// TIA Portal V18 export
TYPE "UserValidationMdz_out"
   STRUCT
      Station : Array[1.."Station_Setup_Const"] of Struct
         Position : Array[1.."Position_Setup_Const"] of Struct
            User_ID : DInt;
            User_SSB : String[8];
            UserName : String[37];
            MsgLogin : String[40];
            AuthorizedByUserMaster_ID : DInt;
            Authentication : Bool;
         END_STRUCT;
      END_STRUCT;
   END_STRUCT;
   // Station[1].Position[1].User_ID := 0;
   // Station[2].Position[1].User_ID := 0;
   // Station[3].Position[1].User_ID := 0;
   // Station[4].Position[1].User_ID := 0;
   // Station[5].Position[1].User_ID := 0;
   // Station[6].Position[1].User_ID := 0;
   // Station[7].Position[1].User_ID := 0;
   // Station[8].Position[1].User_ID := 0;
   // Station[9].Position[1].User_ID := 0;
   // Station[10].Position[1].User_ID := 0;
   // Station[11].Position[1].User_ID := 0;
   // Station[12].Position[1].User_ID := 0;
   // Station[13].Position[1].User_ID := 0;
   // Station[14].Position[1].User_ID := 0;
   // Station[15].Position[1].User_ID := 0;
   // Station[16].Position[1].User_ID := 0;
   // Station[17].Position[1].User_ID := 0;
   // Station[18].Position[1].User_ID := 0;
   // Station[19].Position[1].User_ID := 0;
   // Station[20].Position[1].User_ID := 0;
   // Station[1].Position[1].User_SSB := '';
   // Station[2].Position[1].User_SSB := '';
   // Station[3].Position[1].User_SSB := '';
   // Station[4].Position[1].User_SSB := '';
   // Station[5].Position[1].User_SSB := '';
   // Station[6].Position[1].User_SSB := '';
   // Station[7].Position[1].User_SSB := '';
   // Station[8].Position[1].User_SSB := '';
   // Station[9].Position[1].User_SSB := '';
   // Station[10].Position[1].User_SSB := '';
   // Station[11].Position[1].User_SSB := '';
   // Station[12].Position[1].User_SSB := '';
   // Station[13].Position[1].User_SSB := '';
   // Station[14].Position[1].User_SSB := '';
   // Station[15].Position[1].User_SSB := '';
   // Station[16].Position[1].User_SSB := '';
   // Station[17].Position[1].User_SSB := '';
   // Station[18].Position[1].User_SSB := '';
   // Station[19].Position[1].User_SSB := '';
   // Station[20].Position[1].User_SSB := '';
   // Station[1].Position[1].UserName := '';
   // Station[2].Position[1].UserName := '';
   // Station[3].Position[1].UserName := '';
   // Station[4].Position[1].UserName := '';
   // Station[5].Position[1].UserName := '';
   // Station[6].Position[1].UserName := '';
   // Station[7].Position[1].UserName := '';
   // Station[8].Position[1].UserName := '';
   // Station[9].Position[1].UserName := '';
   // Station[10].Position[1].UserName := '';
   // Station[11].Position[1].UserName := '';
   // Station[12].Position[1].UserName := '';
   // Station[13].Position[1].UserName := '';
   // Station[14].Position[1].UserName := '';
   // Station[15].Position[1].UserName := '';
   // Station[16].Position[1].UserName := '';
   // Station[17].Position[1].UserName := '';
   // Station[18].Position[1].UserName := '';
   // Station[19].Position[1].UserName := '';
   // Station[20].Position[1].UserName := '';
   // Station[1].Position[1].MsgLogin := 'POSTO: 1 NAO POSSUI USUARIO CADASTRADO';
   // Station[2].Position[1].MsgLogin := 'POSTO: 1 NAO POSSUI USUARIO CADASTRADO';
   // Station[3].Position[1].MsgLogin := 'POSTO: 1 NAO POSSUI USUARIO CADASTRADO';
   // Station[4].Position[1].MsgLogin := 'POSTO: 1 NAO POSSUI USUARIO CADASTRADO';
   // Station[5].Position[1].MsgLogin := 'POSTO: 1 NAO POSSUI USUARIO CADASTRADO';
   // Station[6].Position[1].MsgLogin := 'POSTO: 1 NAO POSSUI USUARIO CADASTRADO';
   // Station[7].Position[1].MsgLogin := 'POSTO: 1 NAO POSSUI USUARIO CADASTRADO';
   // Station[8].Position[1].MsgLogin := 'POSTO: 1 NAO POSSUI USUARIO CADASTRADO';
   // Station[9].Position[1].MsgLogin := 'POSTO: 1 NAO POSSUI USUARIO CADASTRADO';
   // Station[10].Position[1].MsgLogin := 'POSTO: 1 NAO POSSUI USUARIO CADASTRADO';
   // Station[11].Position[1].MsgLogin := 'POSTO: 1 NAO POSSUI USUARIO CADASTRADO';
   // Station[12].Position[1].MsgLogin := 'POSTO: 1 NAO POSSUI USUARIO CADASTRADO';
   // Station[13].Position[1].MsgLogin := 'POSTO: 1 NAO POSSUI USUARIO CADASTRADO';
   // Station[14].Position[1].MsgLogin := 'POSTO: 1 NAO POSSUI USUARIO CADASTRADO';
   // Station[15].Position[1].MsgLogin := 'POSTO: 1 NAO POSSUI USUARIO CADASTRADO';
   // Station[16].Position[1].MsgLogin := 'POSTO: 1 NAO POSSUI USUARIO CADASTRADO';
   // Station[17].Position[1].MsgLogin := 'POSTO: 1 NAO POSSUI USUARIO CADASTRADO';
   // Station[18].Position[1].MsgLogin := 'POSTO: 1 NAO POSSUI USUARIO CADASTRADO';
   // Station[19].Position[1].MsgLogin := 'POSTO: 1 NAO POSSUI USUARIO CADASTRADO';
   // Station[20].Position[1].MsgLogin := 'POSTO: 1 NAO POSSUI USUARIO CADASTRADO';
   // Station[1].Position[1].AuthorizedByUserMaster_ID := 0;
   // Station[2].Position[1].AuthorizedByUserMaster_ID := 0;
   // Station[3].Position[1].AuthorizedByUserMaster_ID := 0;
   // Station[4].Position[1].AuthorizedByUserMaster_ID := 0;
   // Station[5].Position[1].AuthorizedByUserMaster_ID := 0;
   // Station[6].Position[1].AuthorizedByUserMaster_ID := 0;
   // Station[7].Position[1].AuthorizedByUserMaster_ID := 0;
   // Station[8].Position[1].AuthorizedByUserMaster_ID := 0;
   // Station[9].Position[1].AuthorizedByUserMaster_ID := 0;
   // Station[10].Position[1].AuthorizedByUserMaster_ID := 0;
   // Station[11].Position[1].AuthorizedByUserMaster_ID := 0;
   // Station[12].Position[1].AuthorizedByUserMaster_ID := 0;
   // Station[13].Position[1].AuthorizedByUserMaster_ID := 0;
   // Station[14].Position[1].AuthorizedByUserMaster_ID := 0;
   // Station[15].Position[1].AuthorizedByUserMaster_ID := 0;
   // Station[16].Position[1].AuthorizedByUserMaster_ID := 0;
   // Station[17].Position[1].AuthorizedByUserMaster_ID := 0;
   // Station[18].Position[1].AuthorizedByUserMaster_ID := 0;
   // Station[19].Position[1].AuthorizedByUserMaster_ID := 0;
   // Station[20].Position[1].AuthorizedByUserMaster_ID := 0;
   // Station[1].Position[1].Authentication := FALSE;
   // Station[2].Position[1].Authentication := FALSE;
   // Station[3].Position[1].Authentication := FALSE;
   // Station[4].Position[1].Authentication := FALSE;
   // Station[5].Position[1].Authentication := FALSE;
   // Station[6].Position[1].Authentication := FALSE;
   // Station[7].Position[1].Authentication := FALSE;
   // Station[8].Position[1].Authentication := FALSE;
   // Station[9].Position[1].Authentication := FALSE;
   // Station[10].Position[1].Authentication := FALSE;
   // Station[11].Position[1].Authentication := FALSE;
   // Station[12].Position[1].Authentication := FALSE;
   // Station[13].Position[1].Authentication := FALSE;
   // Station[14].Position[1].Authentication := FALSE;
   // Station[15].Position[1].Authentication := FALSE;
   // Station[16].Position[1].Authentication := FALSE;
   // Station[17].Position[1].Authentication := FALSE;
   // Station[18].Position[1].Authentication := FALSE;
   // Station[19].Position[1].Authentication := FALSE;
   // Station[20].Position[1].Authentication := FALSE;
END_TYPE
